FUNCTION_BLOCK ManualAutomaticSwitch (* Basic Function Block Type *)
  (* Standard: 61499-2 *)
  (* Version 0.0, 10/19/2026, lizar, Schneider Electric, Template *)
  PACKAGE Main;
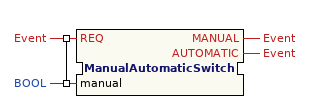
  EVENT_INPUT
    REQ WITH manual; (* Normal Execution Request *)
  END_EVENT
  EVENT_OUTPUT
    MANUAL;
    AUTOMATIC;
  END_EVENT
  VAR_INPUT
    manual : BOOL; (* Input event qualifier *)
  END_VAR
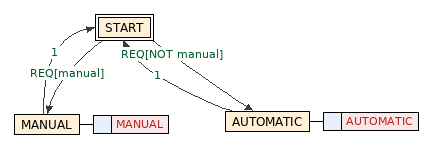
  EC_STATES
    START; (* Initial State *)
    MANUAL : -> MANUAL; (* Normal execution *)
    AUTOMATIC : -> AUTOMATIC;
  END_STATES
  EC_TRANSITIONS
    START TO MANUAL := REQ[manual];
    MANUAL TO START := 1;
    START TO AUTOMATIC := REQ[NOT manual];
    AUTOMATIC TO START := 1;
  END_TRANSITIONS
END_FUNCTION_BLOCK
